(* PLC project probe.project, CODESYS CODESYS V3.5 SP17 Patch 3 *)
(* stored: creationDateTime 2026-10-20T03:54:26.7372477, modificationDateTime 1601-01-01T03:00:00 *)

{attribute 'qualified_only'}
{attribute 'checksumnoinit_override' := '450480064'}
{attribute 'init_related_code' := 'b6ac4937-6a78-4e1e-9458-9c84c4255849'}
VAR_GLOBAL PERSISTENT  (* GVL_ProbeP *)
  {attribute 'order_in_persistent_editor' := '0'}
  xFlag : BOOL;
  {attribute 'order_in_persistent_editor' := '1'}
  rTotal : REAL;
  {attribute 'order_in_persistent_editor' := '2'}
  diHours : DINT;
END_VAR
